Fanuc KAREL source: KA00179.KL

PROGRAM KA00179
%NOLOCKGROUP
VAR
  SRC: ARRAY[4] OF STRING[20]
  DST: ARRAY[4] OF XYZWPR
BEGIN
  DST = SRC
END KA00179
